FUNCTION_BLOCK FB_Cover
VAR_INPUT
	open,
	close,
	enable,
	reset,
	limit_open,
	limit_close: 		BOOL;
END_VAR
VAR_OUTPUT
	error:				BOOL;
	Ready:				BOOL;
	Moving_negative:	BOOL;
	Moving_positive:	BOOL;
	timeout:			BOOL;
END_VAR
VAR
	error_state:	SR;
	//triggers for timeout event for cover
	Cover_timeout:	TON;
	open_timeout: TON := (PT := T#3S);
	close_timeout: TON := (PT := T#3S);
END_VAR


error_state(SET1 := limit_open AND limit_close OR timeout,
			RESET := reset,
			Q1 => error);

IF enable THEN
	Moving_positive := open AND NOT limit_open;
	Moving_negative := close AND NOT limit_close;
END_IF
// A timeout occurs, when we open the cover, and the opened signal does not activate within n seconds.
// The same holds for closing the cover. This should not take longer then 10 seconds
Cover_timeout(IN := NOT (limit_open XOR limit_close) AND (open OR close), PT := T#20S);
open_timeout(IN := open AND limit_open, PT := T#3S);
close_timeout(IN := close AND limit_close, PT := T#3S);
timeout := Cover_timeout.Q OR open_timeout.Q OR close_timeout.Q;

Ready := NOT error;

END_FUNCTION_BLOCK

(* stored: Version 1.1.0.1, ProductVersion 3.1.4024.9
   POU FB_Cover: Id {ff502a3a-f6c6-4825-b511-65bfb253b557}, SpecialFunc None *)
